FUNCTION_BLOCK TestingCycle (* CAT Function Block Type *)
  (* Standard: 61499-2 *)
  (* Version 0.0, 11/20/2026, Schneider Electric, template *)
  PACKAGE Main;
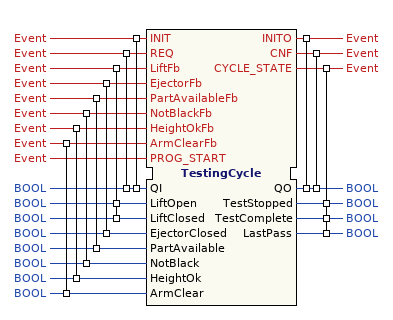
  EVENT_INPUT
    INIT WITH QI; (* Initialization Request *)
    REQ WITH QI; (* Normal Execution Request *)
    LiftFb WITH LiftOpen, LiftClosed;
    EjectorFb WITH EjectorClosed;
    PartAvailableFb WITH PartAvailable;
    NotBlackFb WITH NotBlack;
    HeightOkFb WITH HeightOk;
    ArmClearFb WITH ArmClear;
    PROG_START; (* Programmatic cycle start request *)
  END_EVENT
  EVENT_OUTPUT
    INITO WITH QO; (* Initialization Confirm *)
    CNF WITH QO; (* Execution Confirmation *)
    CYCLE_STATE WITH TestStopped, TestComplete, LastPass; (* Testing cycle state and pass/reject update *)
  END_EVENT
  VAR_INPUT
    QI : BOOL; (* Input event qualifier *)
    LiftOpen : BOOL;
    LiftClosed : BOOL;
    EjectorClosed : BOOL;
    PartAvailable : BOOL;
    NotBlack : BOOL;
    HeightOk : BOOL;
    ArmClear : BOOL;
  END_VAR
  VAR_OUTPUT
    QO : BOOL; (* Output event qualifier *)
    TestStopped : BOOL; (* TRUE when CycleSeq is Stopped *)
    TestComplete : BOOL; (* TRUE when CycleSeq is Completed *)
    LastPass : BOOL; (* TRUE when last cycle took the pass branch (TC10) *)
  END_VAR
  FBS
    CycleSeq : SeqHead(PermStart := TRUE);
    TC1_TakeOver : SeqStep(TransStepId := 2);
    TC2_EnsureBottom : SeqStep(TransStepId := 3);
    TC3_WaitPart : SeqStep(TransStepId := 4);
    TC4_CheckColor : SeqStep(TransStepId := 5);
    TC4_RejectBranch : SeqTransition(TransNextStepId := 11);
    TC5_RaiseLift : SeqStep(TransStepId := 6);
    TC6_CheckHeight : SeqStep(TransStepId := 7);
    TC6_RejectBranch : SeqTransition(TransNextStepId := 11);
    TC7_PassEject : SeqStep(TransStepId := 8);
    TC8_PassRetract : SeqStep(TransStepId := 9);
    TC9_SlideWait : SeqStep(TransStepId := 10);
    TC10_LowerLift : SeqStep(TransStepId := 14);
    TC11_RejectLower : SeqStep(TransStepId := 12);
    TC12_RejectEject : SeqStep(TransStepId := 13);
    TC13_RejectRetract : SeqStep(TransStepId := 14);
    TC14_Finish : SeqStep(TransStepId := 15, Exceeded := TRUE);
    TC_End : SeqTerminate;
    Consts : ANY2ANY_25FC8D56FEEDC9B5(IN1 := TRUE, IN2 := 1, IN3 := 2, IN4 := 0); {SET_ATTRIBUTE(Configuration.GenericFBType.InterfaceParams, Runtime.Standard#CNT:=4;IN${CNT$}:BOOL,INT,INT,INT;OUT${CNT$}:VTQBOOL,VTQINT,VTQINT,VTQINT)}
    OwnerFb : SYMLINKMULTIVARDST_105A0442B8CC61A96(QI := TRUE, NAME1 := 'RES0.Testing.Ejector.sc.progLocal', NAME2 := 'RES0.Testing.AirSlide.sc.progLocal', NAME3 := 'RES0.Testing.Lift.sc.progLocal'); {SET_ATTRIBUTE(Configuration.GenericFBType.InterfaceParams, Runtime.System#I:=3;VALUE${I$}:VTQBOOL,VTQBOOL,VTQBOOL)}
    TakeOverCmd : SYMLINKMULTIVARSRC_105A0442B8CC61A96(QI := TRUE, NAME1 := 'RES0.Testing.Ejector.sc.progLocalSel', NAME2 := 'RES0.Testing.AirSlide.sc.progLocalSel', NAME3 := 'RES0.Testing.Lift.sc.progLocalSel'); {SET_ATTRIBUTE(Configuration.GenericFBType.InterfaceParams, Runtime.System#I:=3;VALUE${I$}:VTQBOOL,VTQBOOL,VTQBOOL)}
    AllLocal : AND_550FE6D62F509EB3(IN3 := TRUE); {SET_ATTRIBUTE(Configuration.GenericFBType.InterfaceParams, Runtime.Standard#CNT:=3;OUT:BOOL)}
    AtBottomReady : AND_550FE6D62F509EB3(IN3 := TRUE); {SET_ATTRIBUTE(Configuration.GenericFBType.InterfaceParams, Runtime.Standard#CNT:=3;OUT:BOOL)}
    IsBlack : NOT_42C76073DCEB1A7A; {SET_ATTRIBUTE(Configuration.GenericFBType.InterfaceParams, Runtime.Standard#CNT:=1;OUT${CNT$}:BOOL)}
    BadHeight : NOT_42C76073DCEB1A7A; {SET_ATTRIBUTE(Configuration.GenericFBType.InterfaceParams, Runtime.Standard#CNT:=1;OUT${CNT$}:BOOL)}
    RaiseLiftCmd : SYMLINKMULTIVARSRC_18556BCA74EA878F1(QI := TRUE, NAME1 := 'RES0.Testing.Lift.sc.lsp'); {SET_ATTRIBUTE(Configuration.GenericFBType.InterfaceParams, Runtime.System#I:=1;VALUE${I$}:VTQINT)}
    LowerLiftCmd : SYMLINKMULTIVARSRC_18556BCA74EA878F1(QI := TRUE, NAME1 := 'RES0.Testing.Lift.sc.lsp'); {SET_ATTRIBUTE(Configuration.GenericFBType.InterfaceParams, Runtime.System#I:=1;VALUE${I$}:VTQINT)}
    ExtendEjectorCmd : SYMLINKMULTIVARSRC_18556BCA74EA878F1(QI := TRUE, NAME1 := 'RES0.Testing.Ejector.sc.lsp'); {SET_ATTRIBUTE(Configuration.GenericFBType.InterfaceParams, Runtime.System#I:=1;VALUE${I$}:VTQINT)}
    RetractEjectorCmd : SYMLINKMULTIVARSRC_18556BCA74EA878F1(QI := TRUE, NAME1 := 'RES0.Testing.Ejector.sc.lsp'); {SET_ATTRIBUTE(Configuration.GenericFBType.InterfaceParams, Runtime.System#I:=1;VALUE${I$}:VTQINT)}
    AirSlideOnCmd : SYMLINKMULTIVARSRC_18556BCA74EA878F1(QI := TRUE, NAME1 := 'RES0.Testing.AirSlide.sc.lsp'); {SET_ATTRIBUTE(Configuration.GenericFBType.InterfaceParams, Runtime.System#I:=1;VALUE${I$}:VTQINT)}
    AirSlideOffCmd : SYMLINKMULTIVARSRC_18556BCA74EA878F1(QI := TRUE, NAME1 := 'RES0.Testing.AirSlide.sc.lsp'); {SET_ATTRIBUTE(Configuration.GenericFBType.InterfaceParams, Runtime.System#I:=1;VALUE${I$}:VTQINT)}
    PassEjectTimer : E_DELAY(DT := T#1s);
    PassEjectLatch : E_SR;
    SlideTimer : E_DELAY(DT := T#2s);
    SlideLatch : E_SR;
    RejEjectTimer : E_DELAY(DT := T#1s);
    RejEjectLatch : E_SR;
    PartAndArmClear : AND_550FE6D62F509EB3(IN3 := TRUE); {SET_ATTRIBUTE(Configuration.GenericFBType.InterfaceParams, Runtime.Standard#CNT:=3;OUT:BOOL)}
    PassResultLatch : E_SR;
  END_FBS
  EVENT_CONNECTIONS
    INIT TO Consts.REQ;
    INIT TO IsBlack.REQ;
    INIT TO BadHeight.REQ;
    Consts.CNF TO CycleSeq.REQ_PERM;
    Consts.CNF TO OwnerFb.INIT;
    Consts.CNF TO TakeOverCmd.INIT;
    Consts.CNF TO RaiseLiftCmd.INIT;
    Consts.CNF TO LowerLiftCmd.INIT;
    Consts.CNF TO ExtendEjectorCmd.INIT;
    Consts.CNF TO RetractEjectorCmd.INIT;
    Consts.CNF TO AirSlideOnCmd.INIT;
    Consts.CNF TO AirSlideOffCmd.INIT;
    TC1_TakeOver.STEP_ENTER TO TakeOverCmd.REQ;
    TakeOverCmd.CNF TO AllLocal.REQ;
    OwnerFb.CNF TO AllLocal.REQ;
    AllLocal.CNF TO TC1_TakeOver.TRANS_REQ;
    TC2_EnsureBottom.STEP_ENTER TO LowerLiftCmd.REQ;
    TC2_EnsureBottom.STEP_ENTER TO RetractEjectorCmd.REQ;
    LowerLiftCmd.CNF TO AtBottomReady.REQ;
    RetractEjectorCmd.CNF TO AtBottomReady.REQ;
    LiftFb TO AtBottomReady.REQ;
    EjectorFb TO AtBottomReady.REQ;
    AtBottomReady.CNF TO TC2_EnsureBottom.TRANS_REQ;
    TC3_WaitPart.STEP_ENTER TO PartAndArmClear.REQ;
    PartAvailableFb TO PartAndArmClear.REQ;
    ArmClearFb TO PartAndArmClear.REQ;
    PartAndArmClear.CNF TO TC3_WaitPart.TRANS_REQ;
    TC4_CheckColor.STEP_ENTER TO TC4_CheckColor.TRANS_REQ;
    NotBlackFb TO TC4_CheckColor.TRANS_REQ;
    TC4_CheckColor.STEP_ENTER TO IsBlack.REQ;
    NotBlackFb TO IsBlack.REQ;
    IsBlack.CNF TO TC4_RejectBranch.TRANS_REQ;
    TC5_RaiseLift.STEP_ENTER TO RaiseLiftCmd.REQ;
    RaiseLiftCmd.CNF TO TC5_RaiseLift.TRANS_REQ;
    LiftFb TO TC5_RaiseLift.TRANS_REQ;
    TC6_CheckHeight.STEP_ENTER TO TC6_CheckHeight.TRANS_REQ;
    HeightOkFb TO TC6_CheckHeight.TRANS_REQ;
    TC6_CheckHeight.STEP_ENTER TO BadHeight.REQ;
    HeightOkFb TO BadHeight.REQ;
    BadHeight.CNF TO TC6_RejectBranch.TRANS_REQ;
    TC7_PassEject.STEP_ENTER TO PassEjectLatch.R;
    TC7_PassEject.STEP_ENTER TO AirSlideOnCmd.REQ;
    TC7_PassEject.STEP_ENTER TO ExtendEjectorCmd.REQ;
    TC7_PassEject.STEP_ENTER TO PassEjectTimer.START;
    PassEjectTimer.EO TO PassEjectLatch.S;
    PassEjectLatch.EO TO TC7_PassEject.TRANS_REQ;
    TC7_PassEject.STEP_LEAVE TO PassEjectTimer.STOP;
    TC7_PassEject.STEP_LEAVE TO PassEjectLatch.R;
    TC8_PassRetract.STEP_ENTER TO RetractEjectorCmd.REQ;
    RetractEjectorCmd.CNF TO TC8_PassRetract.TRANS_REQ;
    EjectorFb TO TC8_PassRetract.TRANS_REQ;
    TC9_SlideWait.STEP_ENTER TO SlideLatch.R;
    TC9_SlideWait.STEP_ENTER TO SlideTimer.START;
    SlideTimer.EO TO SlideLatch.S;
    SlideLatch.EO TO TC9_SlideWait.TRANS_REQ;
    TC9_SlideWait.STEP_LEAVE TO AirSlideOffCmd.REQ;
    TC9_SlideWait.STEP_LEAVE TO SlideTimer.STOP;
    TC9_SlideWait.STEP_LEAVE TO SlideLatch.R;
    TC10_LowerLift.STEP_ENTER TO LowerLiftCmd.REQ;
    LowerLiftCmd.CNF TO TC10_LowerLift.TRANS_REQ;
    LiftFb TO TC10_LowerLift.TRANS_REQ;
    TC11_RejectLower.STEP_ENTER TO LowerLiftCmd.REQ;
    LowerLiftCmd.CNF TO TC11_RejectLower.TRANS_REQ;
    LiftFb TO TC11_RejectLower.TRANS_REQ;
    TC12_RejectEject.STEP_ENTER TO RejEjectLatch.R;
    TC12_RejectEject.STEP_ENTER TO ExtendEjectorCmd.REQ;
    TC12_RejectEject.STEP_ENTER TO RejEjectTimer.START;
    RejEjectTimer.EO TO RejEjectLatch.S;
    RejEjectLatch.EO TO TC12_RejectEject.TRANS_REQ;
    TC12_RejectEject.STEP_LEAVE TO RejEjectTimer.STOP;
    TC12_RejectEject.STEP_LEAVE TO RejEjectLatch.R;
    TC13_RejectRetract.STEP_ENTER TO RetractEjectorCmd.REQ;
    RetractEjectorCmd.CNF TO TC13_RejectRetract.TRANS_REQ;
    EjectorFb TO TC13_RejectRetract.TRANS_REQ;
    TC14_Finish.STEP_ENTER TO TC14_Finish.TRANS_REQ;
    PROG_START TO CycleSeq.START;
    CycleSeq.STATE_IND TO CYCLE_STATE;
    TC1_TakeOver.STEP_ENTER TO PassResultLatch.R;
    TC11_RejectLower.STEP_ENTER TO PassResultLatch.R;
    TC10_LowerLift.STEP_ENTER TO PassResultLatch.S;
  END_CONNECTIONS
  DATA_CONNECTIONS
    Consts.OUT1 TO TakeOverCmd.VALUE1;
    Consts.OUT1 TO TakeOverCmd.VALUE2;
    Consts.OUT1 TO TakeOverCmd.VALUE3;
    Consts.OUT2 TO RaiseLiftCmd.VALUE1;
    Consts.OUT3 TO LowerLiftCmd.VALUE1;
    Consts.OUT2 TO ExtendEjectorCmd.VALUE1;
    Consts.OUT3 TO RetractEjectorCmd.VALUE1;
    Consts.OUT2 TO AirSlideOnCmd.VALUE1;
    Consts.OUT4 TO AirSlideOffCmd.VALUE1;
    OwnerFb.VALUE1 TO AllLocal.IN1;
    OwnerFb.VALUE2 TO AllLocal.IN2;
    AllLocal.OUT TO TC1_TakeOver.Exceeded;
    LiftClosed TO AtBottomReady.IN1;
    EjectorClosed TO AtBottomReady.IN2;
    AtBottomReady.OUT TO TC2_EnsureBottom.Exceeded;
    PartAvailable TO PartAndArmClear.IN1;
    ArmClear TO PartAndArmClear.IN2;
    PartAndArmClear.OUT TO TC3_WaitPart.Exceeded;
    NotBlack TO TC4_CheckColor.Exceeded;
    NotBlack TO IsBlack.IN1;
    IsBlack.OUT1 TO TC4_RejectBranch.Exceeded;
    LiftOpen TO TC5_RaiseLift.Exceeded;
    HeightOk TO TC6_CheckHeight.Exceeded;
    HeightOk TO BadHeight.IN1;
    BadHeight.OUT1 TO TC6_RejectBranch.Exceeded;
    PassEjectLatch.Q TO TC7_PassEject.Exceeded;
    EjectorClosed TO TC8_PassRetract.Exceeded;
    SlideLatch.Q TO TC9_SlideWait.Exceeded;
    LiftClosed TO TC10_LowerLift.Exceeded;
    LiftClosed TO TC11_RejectLower.Exceeded;
    RejEjectLatch.Q TO TC12_RejectEject.Exceeded;
    EjectorClosed TO TC13_RejectRetract.Exceeded;
    CycleSeq.SeqStopped TO TestStopped;
    CycleSeq.SeqComplete TO TestComplete;
    PassResultLatch.Q TO LastPass;
  END_CONNECTIONS
  ADAPTER_CONNECTIONS
    CycleSeq.ISeqChain TO TC1_TakeOver.ISeqChainIn;
    TC1_TakeOver.ISeqChainOut TO TC2_EnsureBottom.ISeqChainIn;
    TC2_EnsureBottom.ISeqChainOut TO TC3_WaitPart.ISeqChainIn;
    TC3_WaitPart.ISeqChainOut TO TC4_CheckColor.ISeqChainIn;
    TC4_CheckColor.ISeqChainOut TO TC5_RaiseLift.ISeqChainIn;
    TC4_CheckColor.ITransChainOut TO TC4_RejectBranch.ITransChainIn;
    TC5_RaiseLift.ISeqChainOut TO TC6_CheckHeight.ISeqChainIn;
    TC6_CheckHeight.ISeqChainOut TO TC7_PassEject.ISeqChainIn;
    TC6_CheckHeight.ITransChainOut TO TC6_RejectBranch.ITransChainIn;
    TC7_PassEject.ISeqChainOut TO TC8_PassRetract.ISeqChainIn;
    TC8_PassRetract.ISeqChainOut TO TC9_SlideWait.ISeqChainIn;
    TC9_SlideWait.ISeqChainOut TO TC10_LowerLift.ISeqChainIn;
    TC10_LowerLift.ISeqChainOut TO TC11_RejectLower.ISeqChainIn;
    TC11_RejectLower.ISeqChainOut TO TC12_RejectEject.ISeqChainIn;
    TC12_RejectEject.ISeqChainOut TO TC13_RejectRetract.ISeqChainIn;
    TC13_RejectRetract.ISeqChainOut TO TC14_Finish.ISeqChainIn;
    TC14_Finish.ISeqChainOut TO TC_End.ISeqChainIn;
  END_CONNECTIONS
END_FUNCTION_BLOCK
